(* IEC 61131-3 sources: stc/testdata/preprocess, 3 files *)

(* ---- define_local.st ---- *)
{DEFINE USE_FEATURE}
PROGRAM Main
VAR
    y : BOOL;
END_VAR
{IF defined(USE_FEATURE)}
    y := TRUE;
{END_IF}
END_PROGRAM

(* ---- error_directive.st ---- *)
{IF defined(VENDOR_BECKHOFF)}
    (* Beckhoff OK *)
{ELSIF defined(VENDOR_SCHNEIDER)}
    (* Schneider OK *)
{ELSE}
    {ERROR "No supported vendor defined. Use --define VENDOR_BECKHOFF or VENDOR_SCHNEIDER"}
{END_IF}

(* ---- vendor_portable.st ---- *)
PROGRAM Main
VAR
    x : INT;
END_VAR
{IF defined(VENDOR_BECKHOFF)}
    x := 1; (* Beckhoff path *)
{ELSIF defined(VENDOR_SCHNEIDER)}
    x := 2; (* Schneider path *)
{ELSE}
    x := 0; (* Generic path *)
{END_IF}
END_PROGRAM
